Universal Robots URScript: T006_mistralai_Mistral-Large-3-675B-Instruct-2512-NVFP4_baseline_rep1_retry1.urscript

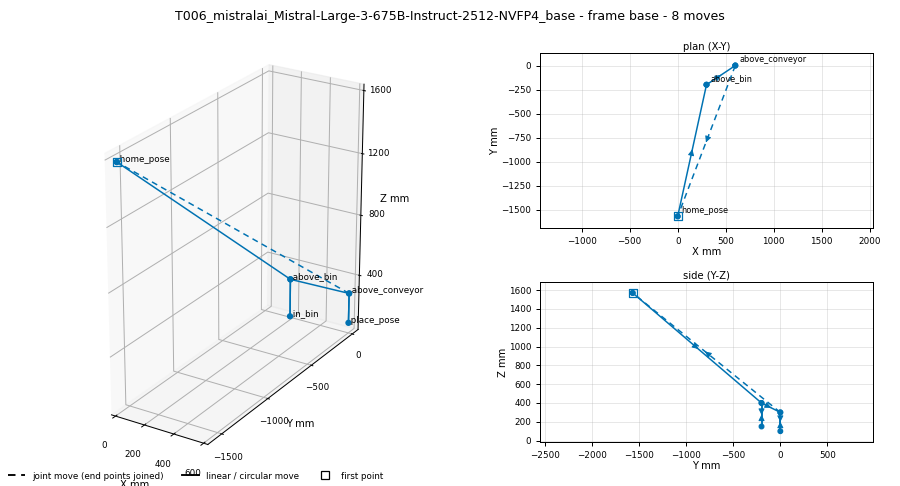
[picture p0: tool path of T006_mistralai_Mistral-Large-3-675B-Instruct-2512-NVFP4_baseline_rep1_retry1.urscript in frame base, 8 of 8 moves have a stored position in this frame; points joined in program order, loops and branches not executed]
# Bin picking with suction - fenced mode (T006)
# Safety parameters
set_analog_inputrange(0, 0)
set_analog_inputrange(1, 0)
set_analog_outputdomain(0, 0)
set_analog_outputdomain(1, 0)
set_tool_voltage(0)
set_runstate_outputs([])
set_payload(2.0)
set_tcp(p[0,0,0.1,0,0,0])

# Safety configuration
conf = { "safety_status": 2, "reduced_mode": False, "operational_mode": 2 }
safetyconf = { "conf": conf }
set_config(safetyconf)

# Watchdog setup
watchdog_min_limit = 0.05
watchdog_max_limit = 0.2
watchdog_input = 0
set_watchdog(watchdog_input, watchdog_min_limit, "watchdog")

# Waypoints
home_pose = p[0.0, -1.5708, 1.5708, -1.5708, -1.5708, 0.0]
above_bin = p[0.3, -0.2, 0.4, 2.221, -2.221, 0.0]
in_bin = p[0.3, -0.2, 0.15, 2.221, -2.221, 0.0]
above_conveyor = p[0.6, 0.0, 0.3, 0.0, 0.0, 0.0]
place_pose = p[0.6, 0.0, 0.1, 0.0, 0.0, 0.0]

# Motion parameters
speed_home = 350.0/1000
speed_above_bin = 350.0/1000
speed_descend = 150.0/1000
speed_lift = 300.0/1000
speed_transit = 380.0/1000
accel = 1.2

# Main program
def main():
    # Enable watchdog
    watchdog()

    # Move to home position
    movej(home_pose, a=accel, v=speed_home)

    # Move above bin
    movel(above_bin, a=accel, v=speed_above_bin)

    # Descend into bin
    movel(in_bin, a=accel, v=speed_descend)

    # Activate suction
    set_tool_digital_out(0, True)
    sleep(0.5)

    # Lift from bin
    movel(above_bin, a=accel, v=speed_lift)

    # Transit to conveyor
    movel(above_conveyor, a=accel, v=speed_transit)

    # Descend to place position
    movel(place_pose, a=accel, v=speed_descend)

    # Release part
    set_tool_digital_out(0, False)
    sleep(0.5)

    # Lift from conveyor
    movel(above_conveyor, a=accel, v=speed_lift)

    # Return to home
    movej(home_pose, a=accel, v=speed_home)

    # Disable watchdog
    watchdog()

end

# Watchdog function
def watchdog():
    if get_configurable_digital_in(0):
        feed_watchdog()
    end
end
